(* Logix 5000 project; controller R400_500_XLS vendor 1 type 14 code 216 rev 31.11; software revision 31.01; part 24 of 32 *)
(* tags used below, declared in another part *)
   Abort1 : DINT;   // Not Used
   CycExcBuffer : UDT_CYCLE;
   Drain_RcvryTnk_with_Sump : DINT;   // 0 = Close Recovery Tank Drain Valve 1 = Open Recovery Tank Drain Valve
   DrainNo : DINT;
   DrnSmp : DINT;
   F1rinse : DINT;   // Not Used
   F2rinse : DINT;   // Not Used
   F3rinse : DINT;   // Not Used
   F4rinse : INT;   // Transition for the conductivity based evalutaion
   FINALRINSE_1 : DINT;   // Final rinse 1 id number
   FINALRINSE_9 : DINT;   // Final rinse 9 id number
   First_PwWshRnseTtr : DINT;
   Last_PwWshRnseTtr : DINT;
   M : DINT[5];   // Memory Bits
   ONS_FC13 : DINT;
   PREWASH_1 : DINT;   // Pre-wash 1 id number
   PREWASH_2 : DINT;   // Pre-wash 2 id number
   PREWASH_3 : DINT;   // Pre-wash 3 id number
   PREWASH_4 : DINT;   // Pre-wash 4 id number
   Rcvry_Tnk_Tmp : REAL;   // Water Temperature of the Heat Recovery Tank
   RINSE_1 : DINT;   // Rinse 1 id number
   RINSE_2 : DINT;   // Rinse 2 id number
   RINSE_3 : DINT;   // Rinse 3 id number
   RINSE_4 : DINT;   // Rinse 4 id number
   RLO : BOOL;   // Logic result
   Run : DINT;
   Shutdown : SINT;   // Shutdown sequence steps
   SumpWaterVolume : DINT;   // Sump Water Volume 0 =Low 1= High
   Tmr : TIMER[107];
   Trt_Drying : SINT;
   Trt_PrWsh : DINT;
   Trt_Rinse : DINT;   // Rinse steps
   Trt_Wsh : DINT;
   WASH_1 : DINT;   // Wash 1 id number
   WASH_2 : DINT;   // Wash 2 id number
   WASH_3 : DINT;   // Wash 3 id number
   WASH_4 : DINT;   // Wash 4 id number
   WASH_5 : DINT;   // Wash 5 id number
   DrainExtensionTime : DINT;
   SumpTemp : REAL;   // Sump temperature in °C
   SumpTempToCool : REAL;   // Sump temperature in °C
   TreatmentPtr : DINT;
   Unit : Hrdwre;   // Unit Configuration
(* MainProgram, continued *)

ROUTINE WSH_22_DRN_SMP_RCVR_TNK   (* ladder *)
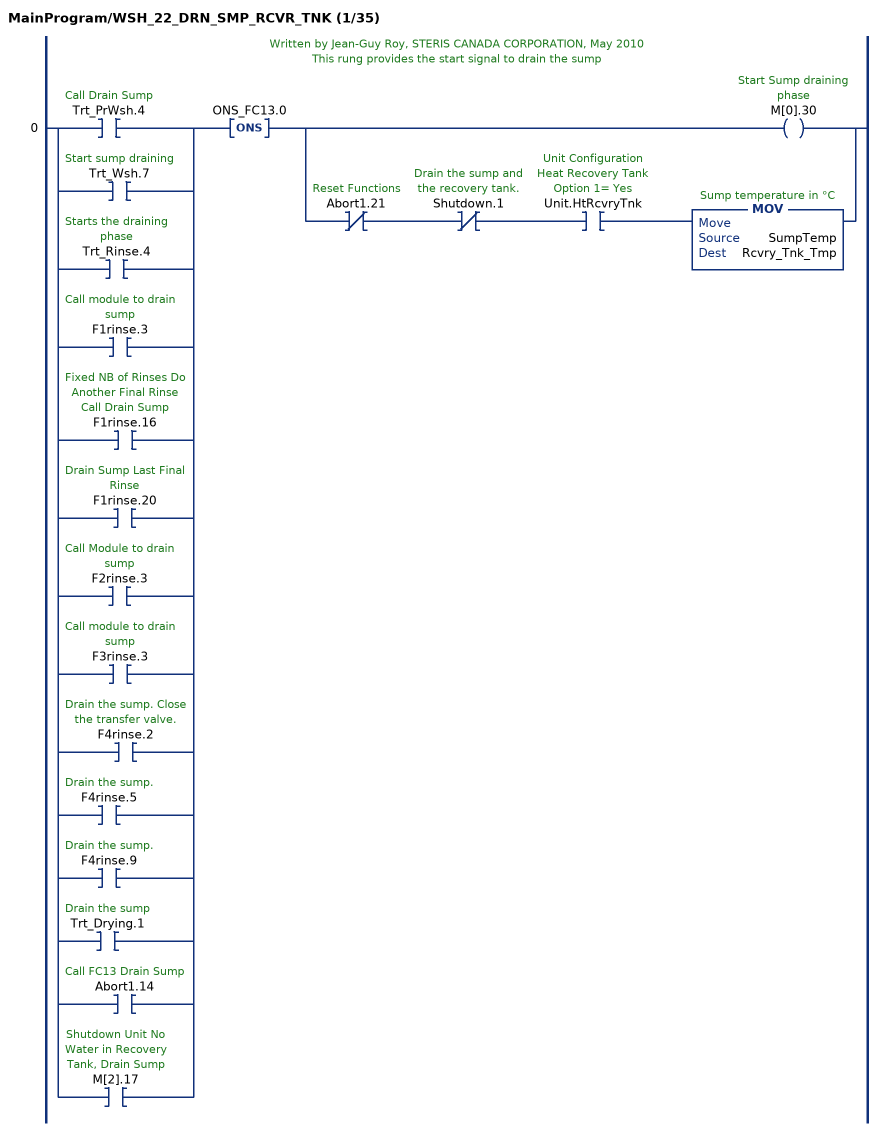
   // Written by Jean-Guy Roy, STERIS CANADA CORPORATION, May 2010
   // This rung provides the start signal to drain the sump
   0: [XIC(Trt_PrWsh.4) ,XIC(Trt_Wsh.7) ,XIC(Trt_Rinse.4) ,XIC(F1rinse.3) ,XIC(F1rinse.16) ,XIC(F1rinse.20) ,XIC(F2rinse.3) ,XIC(F3rinse.3) ,XIC(F4rinse.2) ,XIC(F4rinse.5) ,XIC(F4rinse.9) ,XIC(Trt_Drying.1) ,XIC(Abort1.14) ,XIC(M[2].17) ]ONS(ONS_FC13.0)[OTE(M[0].30) ,XIO(Abort1.21) XIO(Shutdown.1) XIC(Unit.HtRcvryTnk) MOV(SumpTemp,Rcvry_Tnk_Tmp) ];
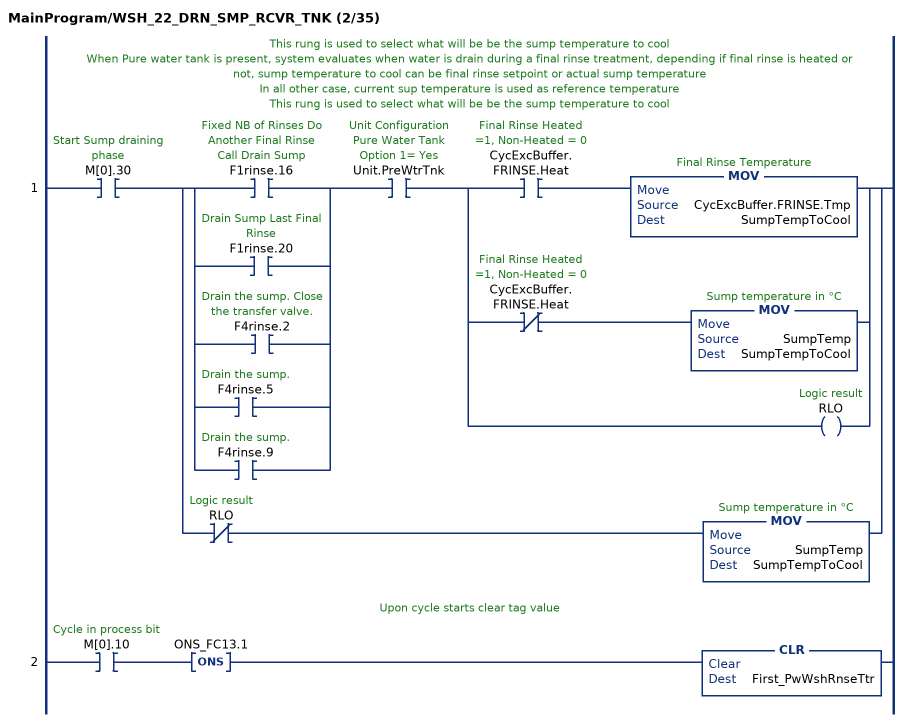
   // This rung is used to select what will be be the sump temperature to cool
   // When Pure water tank is present, system evaluates when water is drain during a final rinse treatment, depending if final rinse is heated or not, sump temperature to cool can be final rinse setpoint or actual sump temperature
   // In all other case, current sup temperature is used as reference temperature
   // This rung is used to select what will be be the sump temperature to cool
   1: XIC(M[0].30)[[XIC(F1rinse.16) ,XIC(F1rinse.20) ,XIC(F4rinse.2) ,XIC(F4rinse.5) ,XIC(F4rinse.9) ] XIC(Unit.PreWtrTnk) [XIC(CycExcBuffer.FRINSE.Heat) MOV(CycExcBuffer.FRINSE.Tmp,SumpTempToCool) ,XIO(CycExcBuffer.FRINSE.Heat) MOV(SumpTemp,SumpTempToCool) ,OTE(RLO) ] ,XIO(RLO) MOV(SumpTemp,SumpTempToCool) ];
   // Upon cycle starts clear tag value
   2: XIC(M[0].10)ONS(ONS_FC13.1)CLR(First_PwWshRnseTtr);
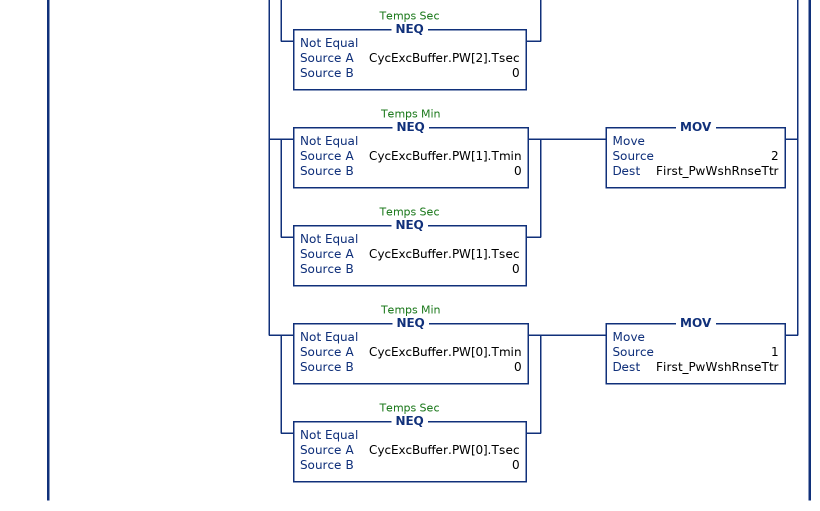
   // This rung checks which Pre-wash, Wash or Rinse treatment is the first treatment of the cycle
   // XLSV10  DGB  2018-09-17 : Added To support New Treatment
   3: XIC(M[0].10)ONS(ONS_FC13.2)[[NEQ(CycExcBuffer.RINSE[3].Tmin,0) ,NEQ(CycExcBuffer.RINSE[3].Tsec,0) ] MOV(13,First_PwWshRnseTtr) ,[NEQ(CycExcBuffer.RINSE[2].Tmin,0) ,NEQ(CycExcBuffer.RINSE[2].Tsec,0) ] MOV(12,First_PwWshRnseTtr) ,[NEQ(CycExcBuffer.RINSE[1].Tmin,0) ,NEQ(CycExcBuffer.RINSE[1].Tsec,0) ] MOV(11,First_PwWshRnseTtr) ,[NEQ(CycExcBuffer.RINSE[0].Tmin,0) ,NEQ(CycExcBuffer.RINSE[0].Tsec,0) ] MOV(10,First_PwWshRnseTtr) ,[NEQ(CycExcBuffer.WSH[4].Tmin,0) ,NEQ(CycExcBuffer.WSH[4].Tsec,0) ] MOV(9,First_PwWshRnseTtr) ,[NEQ(CycExcBuffer.WSH[3].Tmin,0) ,NEQ(CycExcBuffer.WSH[3].Tsec,0) ] MOV(8,First_PwWshRnseTtr) ,[NEQ(CycExcBuffer.WSH[2].Tmin,0) ,NEQ(CycExcBuffer.WSH[2].Tsec,0) ] MOV(7,First_PwWshRnseTtr) ,[NEQ(CycExcBuffer.WSH[1].Tmin,0) ,NEQ(CycExcBuffer.WSH[1].Tsec,0) ] MOV(6,First_PwWshRnseTtr) ,[NEQ(CycExcBuffer.WSH[0].Tmin,0) ,NEQ(CycExcBuffer.WSH[0].Tsec,0) ] MOV(5,First_PwWshRnseTtr) ,[NEQ(CycExcBuffer.PW[3].Tmin,0) ,NEQ(CycExcBuffer.PW[3].Tsec,0) ] MOV(4,First_PwWshRnseTtr) ,[NEQ(CycExcBuffer.PW[2].Tmin,0) ,NEQ(CycExcBuffer.PW[2].Tsec,0) ] MOV(3,First_PwWshRnseTtr) ,[NEQ(CycExcBuffer.PW[1].Tmin,0) ,NEQ(CycExcBuffer.PW[1].Tsec,0) ] MOV(2,First_PwWshRnseTtr) ,[NEQ(CycExcBuffer.PW[0].Tmin,0) ,NEQ(CycExcBuffer.PW[0].Tsec,0) ] MOV(1,First_PwWshRnseTtr) ];
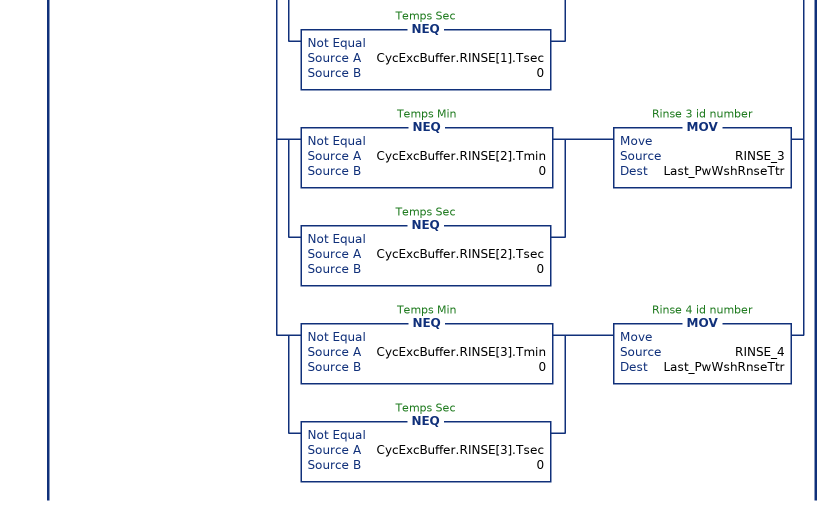
   // This rung detect which recirculated treatment is the last treatment of the cycle
   // XLSV10  DGB  2018-09-07 : Modified to support Added Treatments
   4: XIC(M[0].10)ONS(ONS_FC13.10)[[NEQ(CycExcBuffer.PW[0].Tmin,0) ,NEQ(CycExcBuffer.PW[0].Tsec,0) ] MOV(PREWASH_1,Last_PwWshRnseTtr) ,[NEQ(CycExcBuffer.PW[1].Tmin,0) ,NEQ(CycExcBuffer.PW[1].Tsec,0) ] MOV(PREWASH_2,Last_PwWshRnseTtr) ,[NEQ(CycExcBuffer.PW[2].Tmin,0) ,NEQ(CycExcBuffer.PW[2].Tsec,0) ] MOV(PREWASH_3,Last_PwWshRnseTtr) ,[NEQ(CycExcBuffer.PW[3].Tmin,0) ,NEQ(CycExcBuffer.PW[3].Tsec,0) ] MOV(PREWASH_4,Last_PwWshRnseTtr) ,[NEQ(CycExcBuffer.WSH[0].Tmin,0) ,NEQ(CycExcBuffer.WSH[0].Tsec,0) ] MOV(WASH_1,Last_PwWshRnseTtr) ,[NEQ(CycExcBuffer.WSH[1].Tmin,0) ,NEQ(CycExcBuffer.WSH[1].Tsec,0) ] MOV(WASH_2,Last_PwWshRnseTtr) ,[NEQ(CycExcBuffer.WSH[2].Tmin,0) ,NEQ(CycExcBuffer.WSH[2].Tsec,0) ] MOV(WASH_3,Last_PwWshRnseTtr) ,[NEQ(CycExcBuffer.WSH[3].Tmin,0) ,NEQ(CycExcBuffer.WSH[3].Tsec,0) ] MOV(WASH_4,Last_PwWshRnseTtr) ,[NEQ(CycExcBuffer.WSH[4].Tmin,0) ,NEQ(CycExcBuffer.WSH[4].Tsec,0) ] MOV(WASH_5,Last_PwWshRnseTtr) ,[NEQ(CycExcBuffer.RINSE[0].Tmin,0) ,NEQ(CycExcBuffer.RINSE[0].Tsec,0) ] MOV(RINSE_1,Last_PwWshRnseTtr) ,[NEQ(CycExcBuffer.RINSE[1].Tmin,0) ,NEQ(CycExcBuffer.RINSE[1].Tsec,0) ] MOV(RINSE_2,Last_PwWshRnseTtr) ,[NEQ(CycExcBuffer.RINSE[2].Tmin,0) ,NEQ(CycExcBuffer.RINSE[2].Tsec,0) ] MOV(RINSE_3,Last_PwWshRnseTtr) ,[NEQ(CycExcBuffer.RINSE[3].Tmin,0) ,NEQ(CycExcBuffer.RINSE[3].Tsec,0) ] MOV(RINSE_4,Last_PwWshRnseTtr) ];
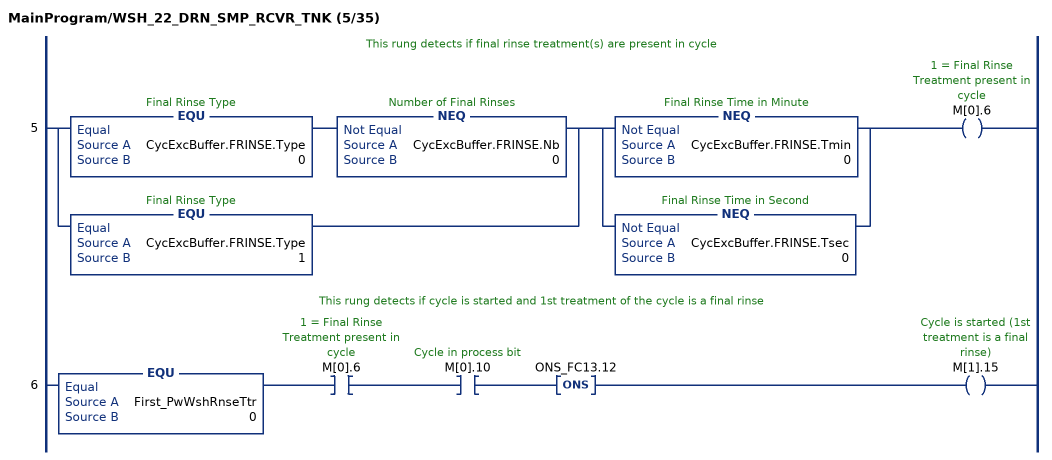
   // This rung detects if final rinse treatment(s) are present in cycle
   5: [EQU(CycExcBuffer.FRINSE.Type,0) NEQ(CycExcBuffer.FRINSE.Nb,0) ,EQU(CycExcBuffer.FRINSE.Type,1) ][NEQ(CycExcBuffer.FRINSE.Tmin,0) ,NEQ(CycExcBuffer.FRINSE.Tsec,0) ]OTE(M[0].6);
   // This rung detects if cycle is started and 1st treatment of the cycle is a final rinse
   6: EQU(First_PwWshRnseTtr,0)XIC(M[0].6)XIC(M[0].10)ONS(ONS_FC13.12)OTE(M[1].15);
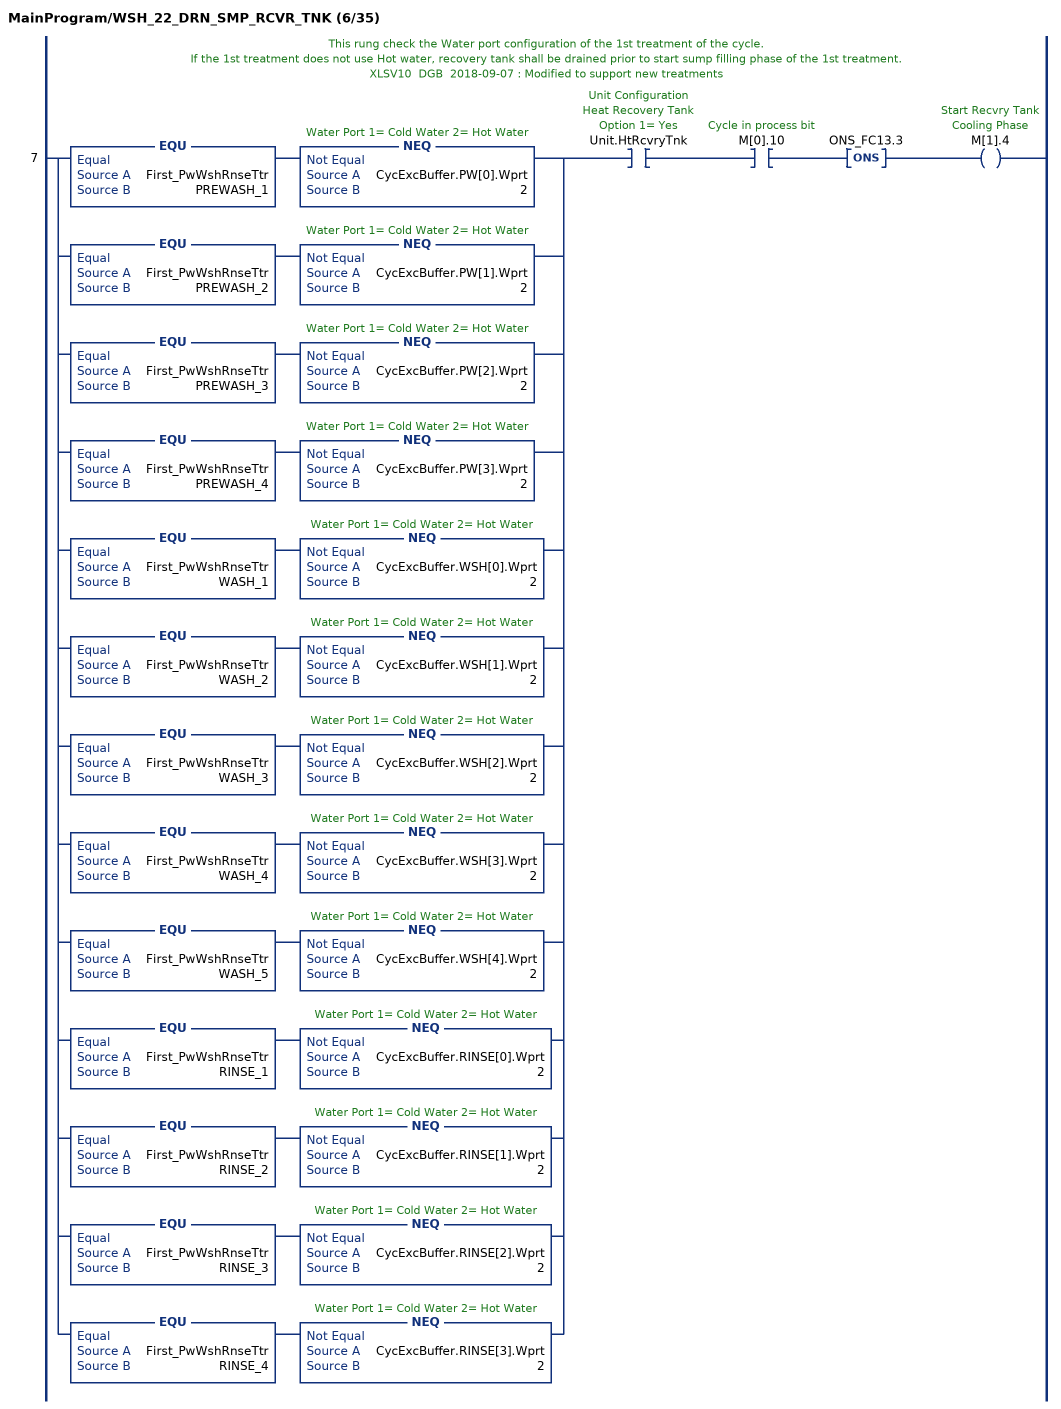
   // This rung check the Water port configuration of the 1st treatment of the cycle.
   // If the 1st treatment does not use Hot water, recovery tank shall be drained prior to start sump filling phase of the 1st treatment.
   // XLSV10  DGB  2018-09-07 : Modified to support new treatments
   7: [EQU(First_PwWshRnseTtr,PREWASH_1) NEQ(CycExcBuffer.PW[0].Wprt,2) ,EQU(First_PwWshRnseTtr,PREWASH_2) NEQ(CycExcBuffer.PW[1].Wprt,2) ,EQU(First_PwWshRnseTtr,PREWASH_3) NEQ(CycExcBuffer.PW[2].Wprt,2) ,EQU(First_PwWshRnseTtr,PREWASH_4) NEQ(CycExcBuffer.PW[3].Wprt,2) ,EQU(First_PwWshRnseTtr,WASH_1) NEQ(CycExcBuffer.WSH[0].Wprt,2) ,EQU(First_PwWshRnseTtr,WASH_2) NEQ(CycExcBuffer.WSH[1].Wprt,2) ,EQU(First_PwWshRnseTtr,WASH_3) NEQ(CycExcBuffer.WSH[2].Wprt,2) ,EQU(First_PwWshRnseTtr,WASH_4) NEQ(CycExcBuffer.WSH[3].Wprt,2) ,EQU(First_PwWshRnseTtr,WASH_5) NEQ(CycExcBuffer.WSH[4].Wprt,2) ,EQU(First_PwWshRnseTtr,RINSE_1) NEQ(CycExcBuffer.RINSE[0].Wprt,2) ,EQU(First_PwWshRnseTtr,RINSE_2) NEQ(CycExcBuffer.RINSE[1].Wprt,2) ,EQU(First_PwWshRnseTtr,RINSE_3) NEQ(CycExcBuffer.RINSE[2].Wprt,2) ,EQU(First_PwWshRnseTtr,RINSE_4) NEQ(CycExcBuffer.RINSE[3].Wprt,2) ]XIC(Unit.HtRcvryTnk)XIC(M[0].10)ONS(ONS_FC13.3)OTE(M[1].4);
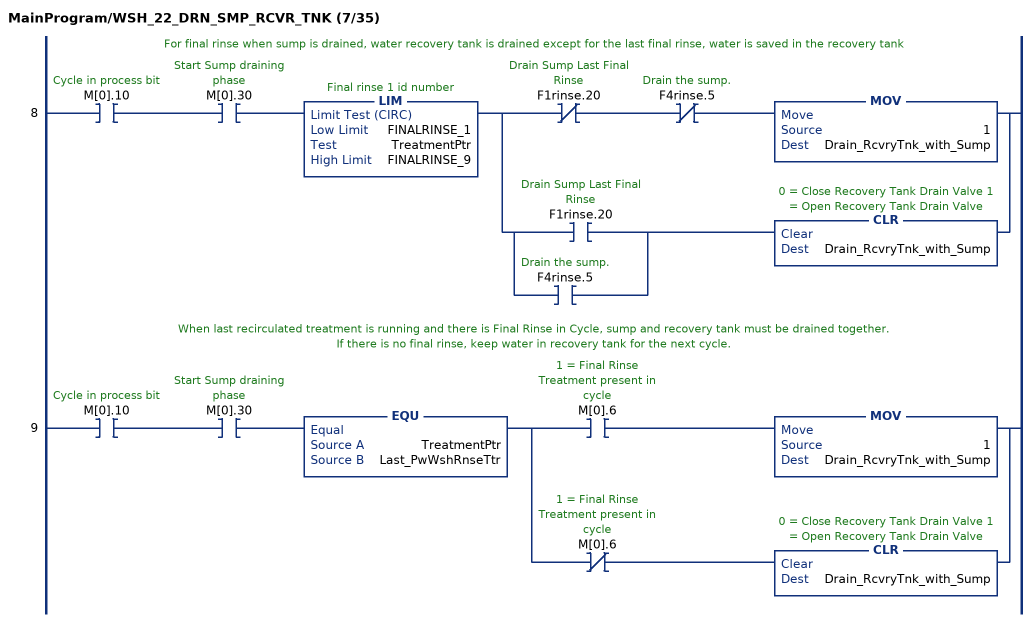
   // For final rinse when sump is drained, water recovery tank is drained except for the last final rinse, water is saved in the recovery tank
   8: XIC(M[0].10)XIC(M[0].30)LIM(FINALRINSE_1,TreatmentPtr,FINALRINSE_9)[XIO(F1rinse.20) XIO(F4rinse.5) MOV(1,Drain_RcvryTnk_with_Sump) ,[XIC(F1rinse.20) ,XIC(F4rinse.5) ] CLR(Drain_RcvryTnk_with_Sump) ];
   // When last recirculated treatment is running and there is Final Rinse in Cycle, sump and recovery tank must be drained together.
   // If there is no final rinse, keep water in recovery tank for the next cycle.
   9: XIC(M[0].10)XIC(M[0].30)EQU(TreatmentPtr,Last_PwWshRnseTtr)[XIC(M[0].6) MOV(1,Drain_RcvryTnk_with_Sump) ,XIO(M[0].6) CLR(Drain_RcvryTnk_with_Sump) ];
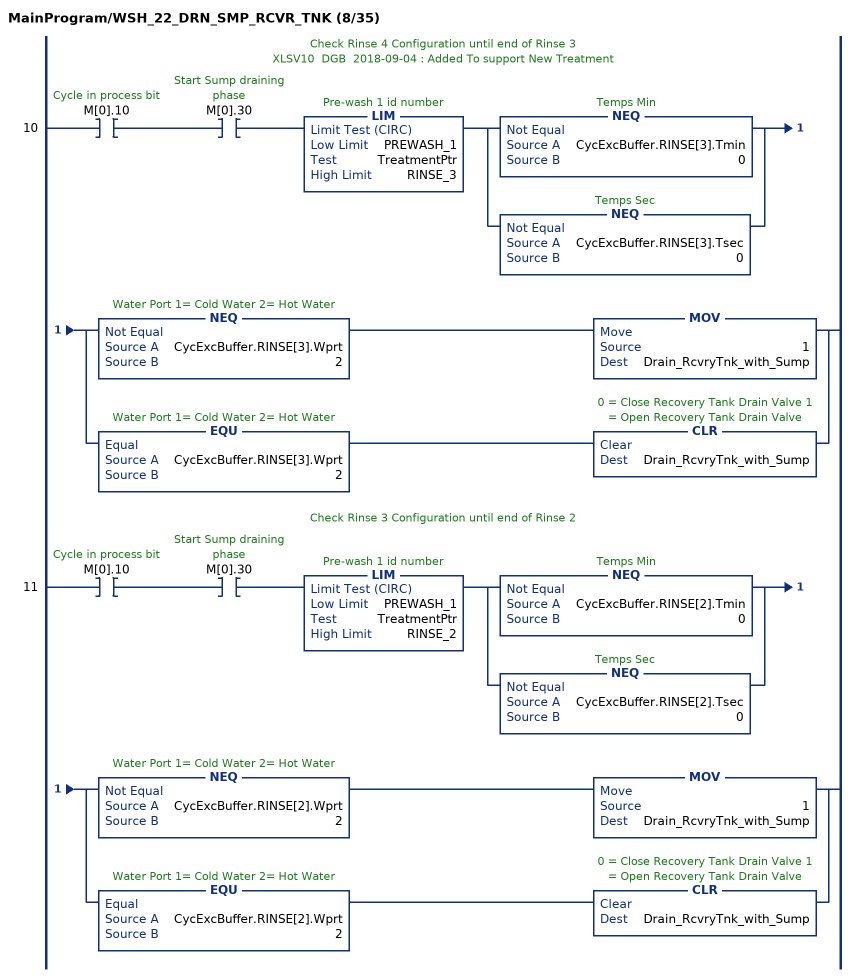
   // Check Rinse 4 Configuration until end of Rinse 3
   // XLSV10  DGB  2018-09-04 : Added To support New Treatment
   10: XIC(M[0].10)XIC(M[0].30)LIM(PREWASH_1,TreatmentPtr,RINSE_3)[NEQ(CycExcBuffer.RINSE[3].Tmin,0) ,NEQ(CycExcBuffer.RINSE[3].Tsec,0) ][NEQ(CycExcBuffer.RINSE[3].Wprt,2) MOV(1,Drain_RcvryTnk_with_Sump) ,EQU(CycExcBuffer.RINSE[3].Wprt,2) CLR(Drain_RcvryTnk_with_Sump) ];
   // Check Rinse 3 Configuration until end of Rinse 2
   11: XIC(M[0].10)XIC(M[0].30)LIM(PREWASH_1,TreatmentPtr,RINSE_2)[NEQ(CycExcBuffer.RINSE[2].Tmin,0) ,NEQ(CycExcBuffer.RINSE[2].Tsec,0) ][NEQ(CycExcBuffer.RINSE[2].Wprt,2) MOV(1,Drain_RcvryTnk_with_Sump) ,EQU(CycExcBuffer.RINSE[2].Wprt,2) CLR(Drain_RcvryTnk_with_Sump) ];
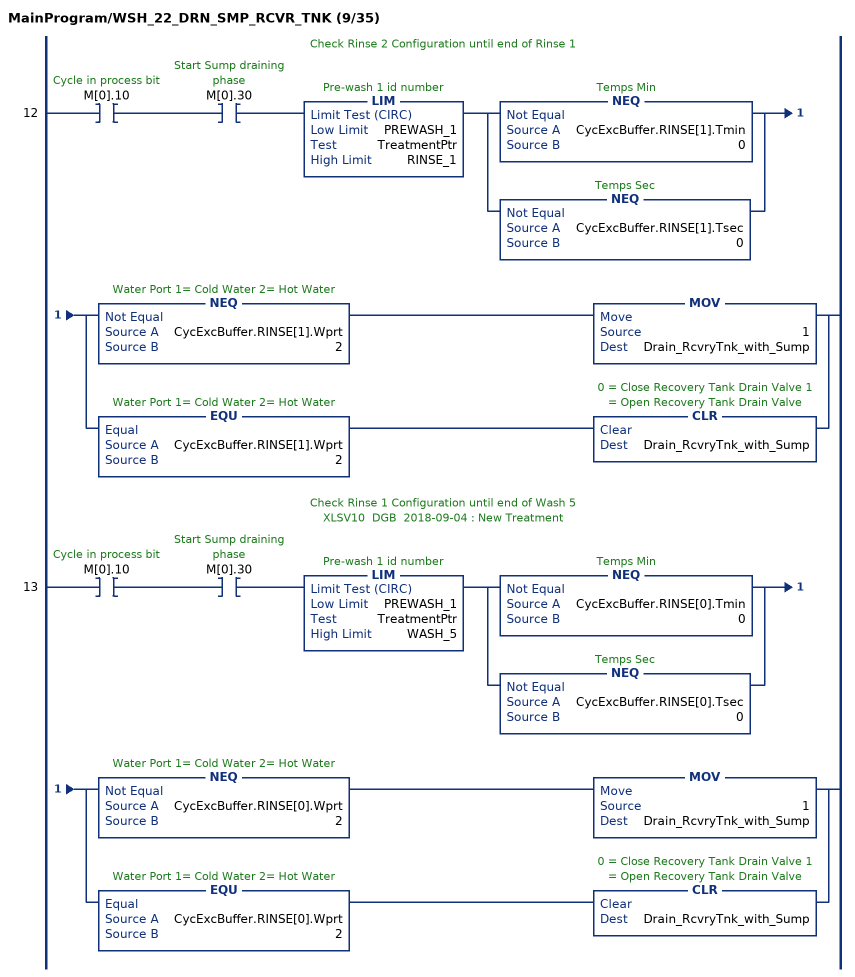
   // Check Rinse 2 Configuration until end of Rinse 1
   12: XIC(M[0].10)XIC(M[0].30)LIM(PREWASH_1,TreatmentPtr,RINSE_1)[NEQ(CycExcBuffer.RINSE[1].Tmin,0) ,NEQ(CycExcBuffer.RINSE[1].Tsec,0) ][NEQ(CycExcBuffer.RINSE[1].Wprt,2) MOV(1,Drain_RcvryTnk_with_Sump) ,EQU(CycExcBuffer.RINSE[1].Wprt,2) CLR(Drain_RcvryTnk_with_Sump) ];
   // Check Rinse 1 Configuration until end of Wash 5
   // XLSV10  DGB  2018-09-04 : New Treatment
   13: XIC(M[0].10)XIC(M[0].30)LIM(PREWASH_1,TreatmentPtr,WASH_5)[NEQ(CycExcBuffer.RINSE[0].Tmin,0) ,NEQ(CycExcBuffer.RINSE[0].Tsec,0) ][NEQ(CycExcBuffer.RINSE[0].Wprt,2) MOV(1,Drain_RcvryTnk_with_Sump) ,EQU(CycExcBuffer.RINSE[0].Wprt,2) CLR(Drain_RcvryTnk_with_Sump) ];
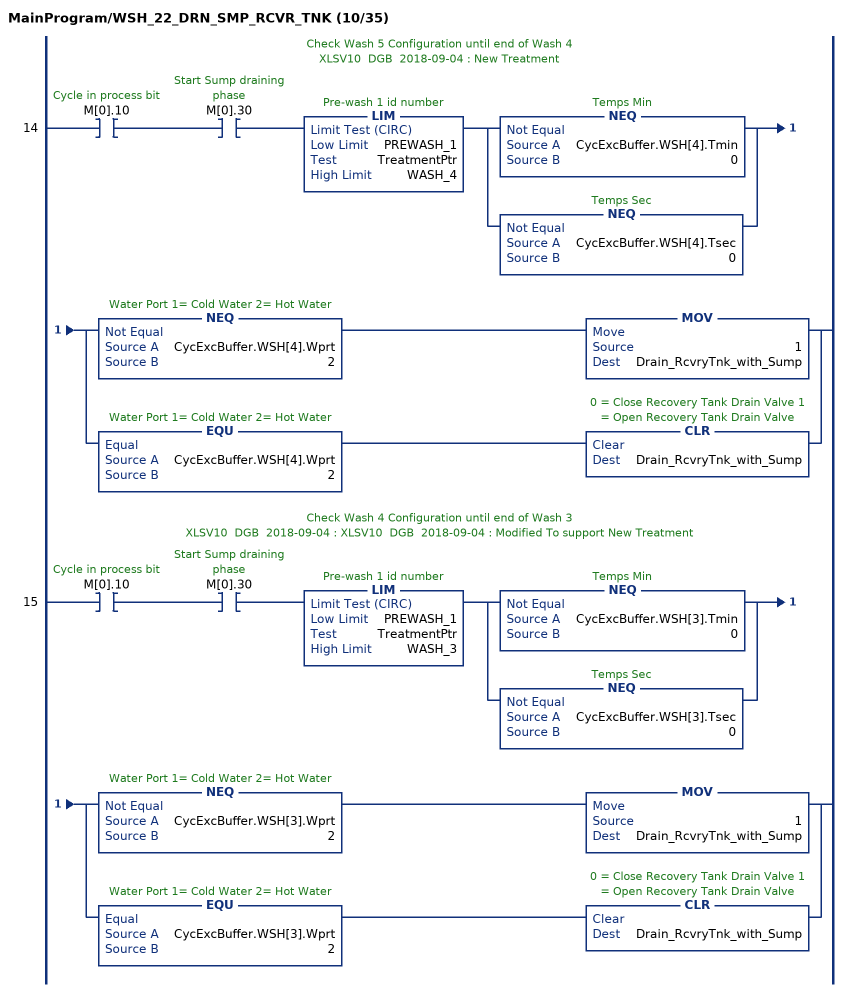
   // Check Wash 5 Configuration until end of Wash 4
   // XLSV10  DGB  2018-09-04 : New Treatment
   14: XIC(M[0].10)XIC(M[0].30)LIM(PREWASH_1,TreatmentPtr,WASH_4)[NEQ(CycExcBuffer.WSH[4].Tmin,0) ,NEQ(CycExcBuffer.WSH[4].Tsec,0) ][NEQ(CycExcBuffer.WSH[4].Wprt,2) MOV(1,Drain_RcvryTnk_with_Sump) ,EQU(CycExcBuffer.WSH[4].Wprt,2) CLR(Drain_RcvryTnk_with_Sump) ];
   // Check Wash 4 Configuration until end of Wash 3
   // XLSV10  DGB  2018-09-04 : XLSV10  DGB  2018-09-04 : Modified To support New Treatment
   15: XIC(M[0].10)XIC(M[0].30)LIM(PREWASH_1,TreatmentPtr,WASH_3)[NEQ(CycExcBuffer.WSH[3].Tmin,0) ,NEQ(CycExcBuffer.WSH[3].Tsec,0) ][NEQ(CycExcBuffer.WSH[3].Wprt,2) MOV(1,Drain_RcvryTnk_with_Sump) ,EQU(CycExcBuffer.WSH[3].Wprt,2) CLR(Drain_RcvryTnk_with_Sump) ];
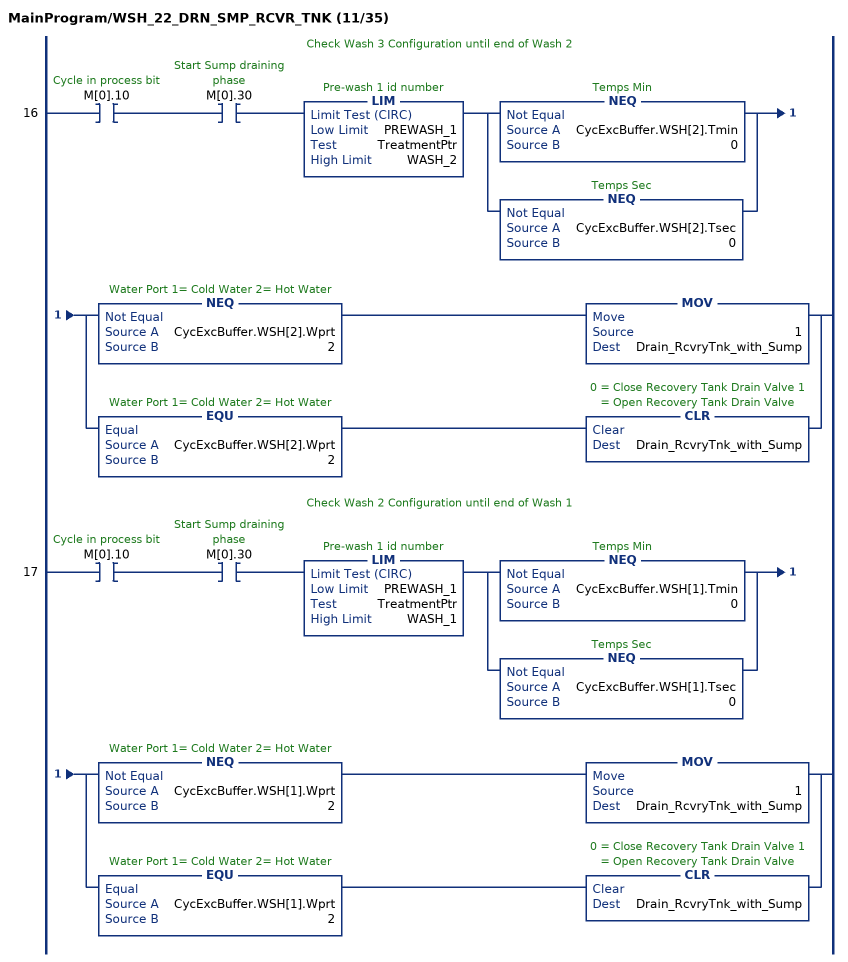
   // Check Wash 3 Configuration until end of Wash 2
   16: XIC(M[0].10)XIC(M[0].30)LIM(PREWASH_1,TreatmentPtr,WASH_2)[NEQ(CycExcBuffer.WSH[2].Tmin,0) ,NEQ(CycExcBuffer.WSH[2].Tsec,0) ][NEQ(CycExcBuffer.WSH[2].Wprt,2) MOV(1,Drain_RcvryTnk_with_Sump) ,EQU(CycExcBuffer.WSH[2].Wprt,2) CLR(Drain_RcvryTnk_with_Sump) ];
   // Check Wash 2 Configuration until end of Wash 1
   17: XIC(M[0].10)XIC(M[0].30)LIM(PREWASH_1,TreatmentPtr,WASH_1)[NEQ(CycExcBuffer.WSH[1].Tmin,0) ,NEQ(CycExcBuffer.WSH[1].Tsec,0) ][NEQ(CycExcBuffer.WSH[1].Wprt,2) MOV(1,Drain_RcvryTnk_with_Sump) ,EQU(CycExcBuffer.WSH[1].Wprt,2) CLR(Drain_RcvryTnk_with_Sump) ];
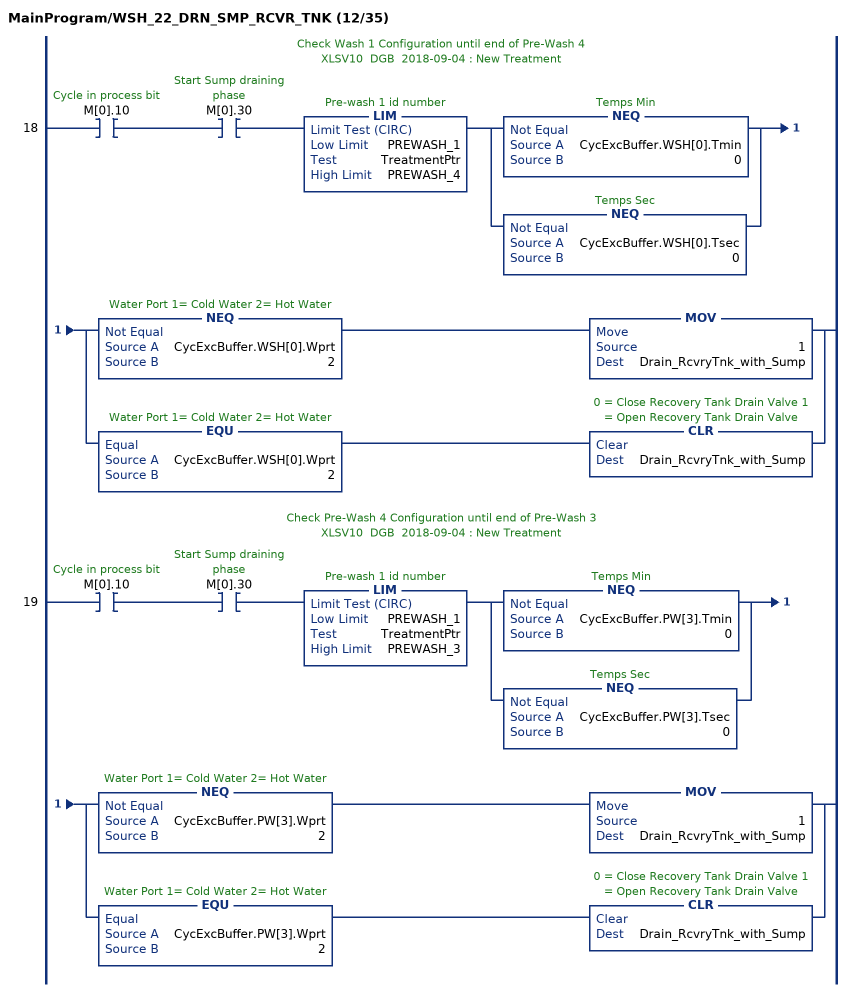
   // Check Wash 1 Configuration until end of Pre-Wash 4
   // XLSV10  DGB  2018-09-04 : New Treatment
   18: XIC(M[0].10)XIC(M[0].30)LIM(PREWASH_1,TreatmentPtr,PREWASH_4)[NEQ(CycExcBuffer.WSH[0].Tmin,0) ,NEQ(CycExcBuffer.WSH[0].Tsec,0) ][NEQ(CycExcBuffer.WSH[0].Wprt,2) MOV(1,Drain_RcvryTnk_with_Sump) ,EQU(CycExcBuffer.WSH[0].Wprt,2) CLR(Drain_RcvryTnk_with_Sump) ];
   // Check Pre-Wash 4 Configuration until end of Pre-Wash 3
   // XLSV10  DGB  2018-09-04 : New Treatment
   19: XIC(M[0].10)XIC(M[0].30)LIM(PREWASH_1,TreatmentPtr,PREWASH_3)[NEQ(CycExcBuffer.PW[3].Tmin,0) ,NEQ(CycExcBuffer.PW[3].Tsec,0) ][NEQ(CycExcBuffer.PW[3].Wprt,2) MOV(1,Drain_RcvryTnk_with_Sump) ,EQU(CycExcBuffer.PW[3].Wprt,2) CLR(Drain_RcvryTnk_with_Sump) ];
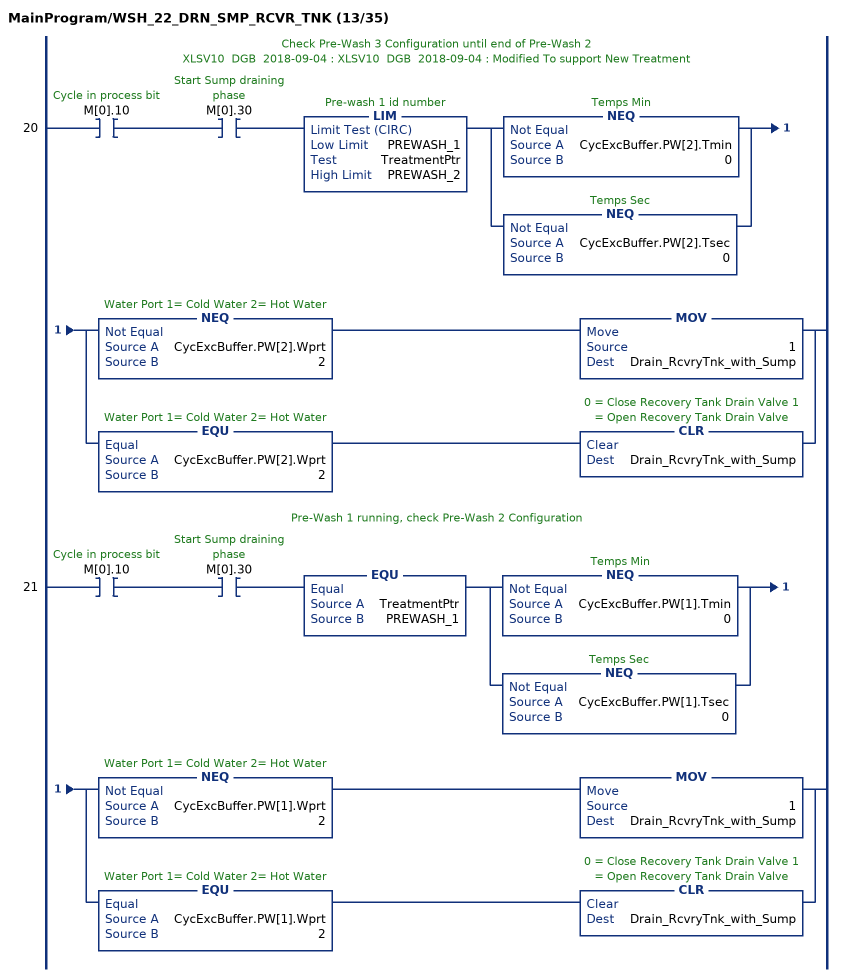
   // Check Pre-Wash 3 Configuration until end of Pre-Wash 2
   // XLSV10  DGB  2018-09-04 : XLSV10  DGB  2018-09-04 : Modified To support New Treatment
   20: XIC(M[0].10)XIC(M[0].30)LIM(PREWASH_1,TreatmentPtr,PREWASH_2)[NEQ(CycExcBuffer.PW[2].Tmin,0) ,NEQ(CycExcBuffer.PW[2].Tsec,0) ][NEQ(CycExcBuffer.PW[2].Wprt,2) MOV(1,Drain_RcvryTnk_with_Sump) ,EQU(CycExcBuffer.PW[2].Wprt,2) CLR(Drain_RcvryTnk_with_Sump) ];
   // Pre-Wash 1 running, check Pre-Wash 2 Configuration
   21: XIC(M[0].10)XIC(M[0].30)EQU(TreatmentPtr,PREWASH_1)[NEQ(CycExcBuffer.PW[1].Tmin,0) ,NEQ(CycExcBuffer.PW[1].Tsec,0) ][NEQ(CycExcBuffer.PW[1].Wprt,2) MOV(1,Drain_RcvryTnk_with_Sump) ,EQU(CycExcBuffer.PW[1].Wprt,2) CLR(Drain_RcvryTnk_with_Sump) ];
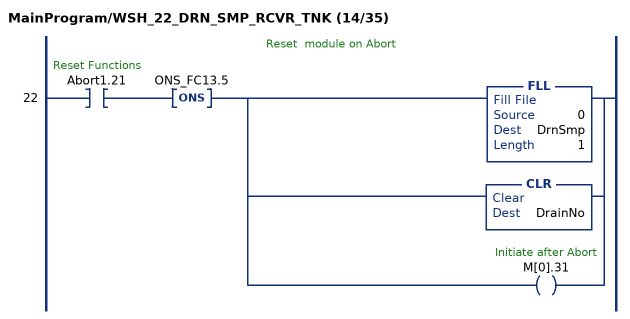
   // Reset  module on Abort
   22: XIC(Abort1.21)ONS(ONS_FC13.5)[FLL(0,DrnSmp,1) ,CLR(DrainNo) ,OTE(M[0].31) ];
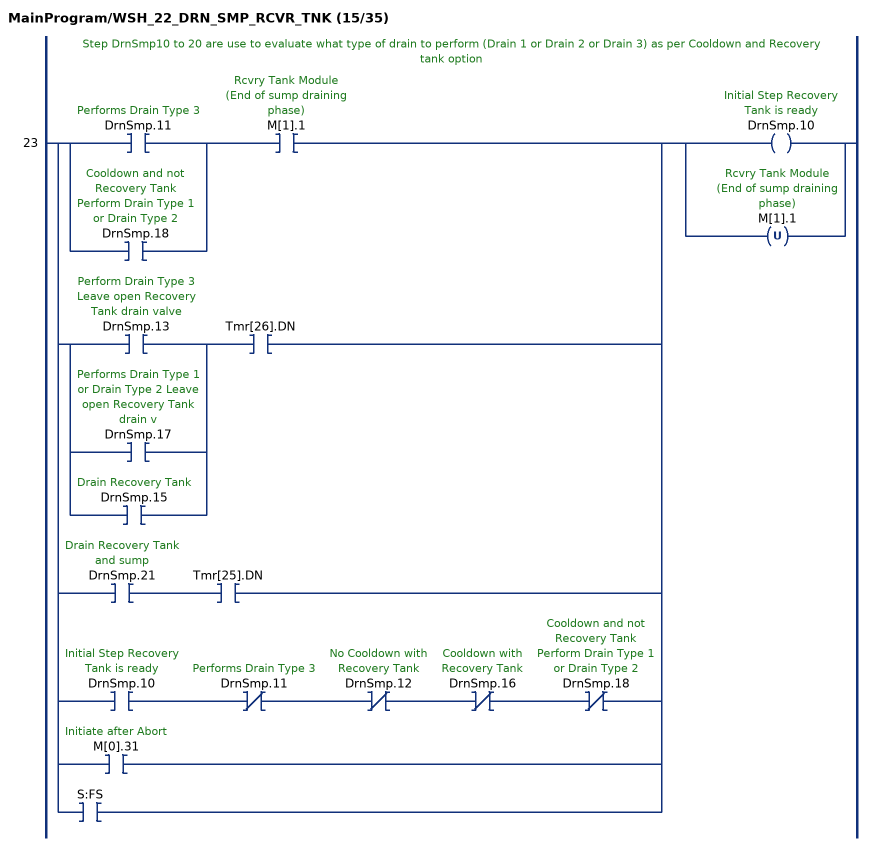
   // Step DrnSmp10 to 20 are use to evaluate what type of drain to perform (Drain 1 or Drain 2 or Drain 3) as per Cooldown and Recovery tank option
   23: [[[XIC(DrnSmp.11) ,XIC(DrnSmp.18) ] XIC(M[1].1) ,[XIC(DrnSmp.13) ,XIC(DrnSmp.17) ,XIC(DrnSmp.15) ] XIC(Tmr[26].DN) ,XIC(DrnSmp.21) XIC(Tmr[25].DN) ] ,XIC(DrnSmp.10) XIO(DrnSmp.11) XIO(DrnSmp.12) XIO(DrnSmp.16) XIO(DrnSmp.18) ,XIC(M[0].31) ,XIC(S:FS) ][OTE(DrnSmp.10) ,OTU(M[1].1) ];
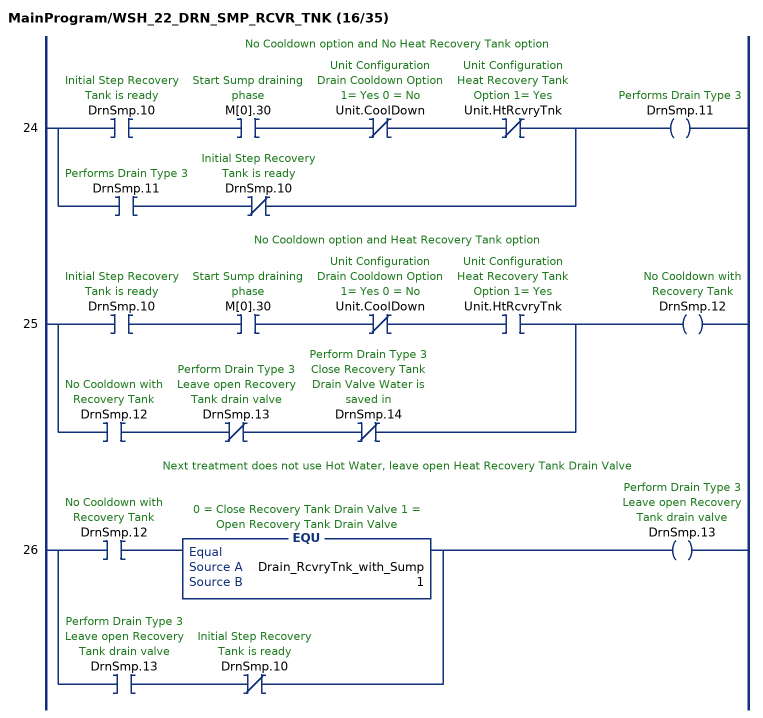
   // No Cooldown option and No Heat Recovery Tank option
   24: [XIC(DrnSmp.10) XIC(M[0].30) XIO(Unit.CoolDown) XIO(Unit.HtRcvryTnk) ,XIC(DrnSmp.11) XIO(DrnSmp.10) ]OTE(DrnSmp.11);
   // No Cooldown option and Heat Recovery Tank option
   25: [XIC(DrnSmp.10) XIC(M[0].30) XIO(Unit.CoolDown) XIC(Unit.HtRcvryTnk) ,XIC(DrnSmp.12) XIO(DrnSmp.13) XIO(DrnSmp.14) ]OTE(DrnSmp.12);
   // Next treatment does not use Hot Water, leave open Heat Recovery Tank Drain Valve
   26: [XIC(DrnSmp.12) EQU(Drain_RcvryTnk_with_Sump,1) ,XIC(DrnSmp.13) XIO(DrnSmp.10) ]OTE(DrnSmp.13);
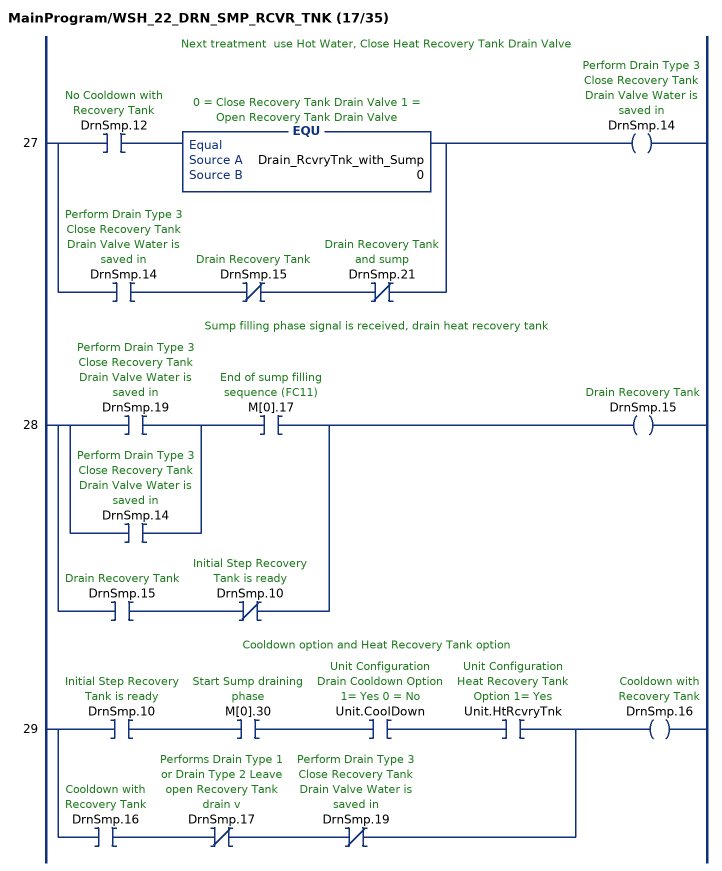
   // Next treatment  use Hot Water, Close Heat Recovery Tank Drain Valve
   27: [XIC(DrnSmp.12) EQU(Drain_RcvryTnk_with_Sump,0) ,XIC(DrnSmp.14) XIO(DrnSmp.15) XIO(DrnSmp.21) ]OTE(DrnSmp.14);
   // Sump filling phase signal is received, drain heat recovery tank
   28: [[XIC(DrnSmp.19) ,XIC(DrnSmp.14) ] XIC(M[0].17) ,XIC(DrnSmp.15) XIO(DrnSmp.10) ]OTE(DrnSmp.15);
   // Cooldown option and Heat Recovery Tank option
   29: [XIC(DrnSmp.10) XIC(M[0].30) XIC(Unit.CoolDown) XIC(Unit.HtRcvryTnk) ,XIC(DrnSmp.16) XIO(DrnSmp.17) XIO(DrnSmp.19) ]OTE(DrnSmp.16);
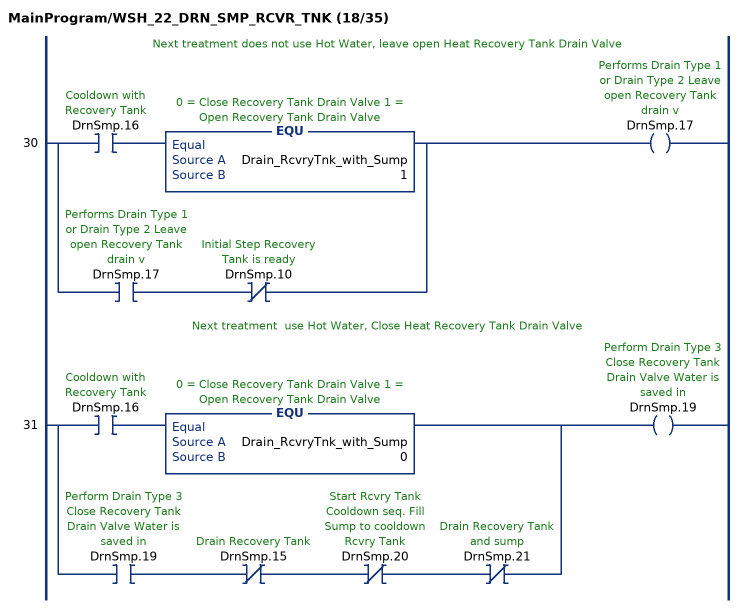
   // Next treatment does not use Hot Water, leave open Heat Recovery Tank Drain Valve
   30: [XIC(DrnSmp.16) EQU(Drain_RcvryTnk_with_Sump,1) ,XIC(DrnSmp.17) XIO(DrnSmp.10) ]OTE(DrnSmp.17);
   // Next treatment  use Hot Water, Close Heat Recovery Tank Drain Valve
   31: [XIC(DrnSmp.16) EQU(Drain_RcvryTnk_with_Sump,0) ,XIC(DrnSmp.19) XIO(DrnSmp.15) XIO(DrnSmp.20) XIO(DrnSmp.21) ]OTE(DrnSmp.19);
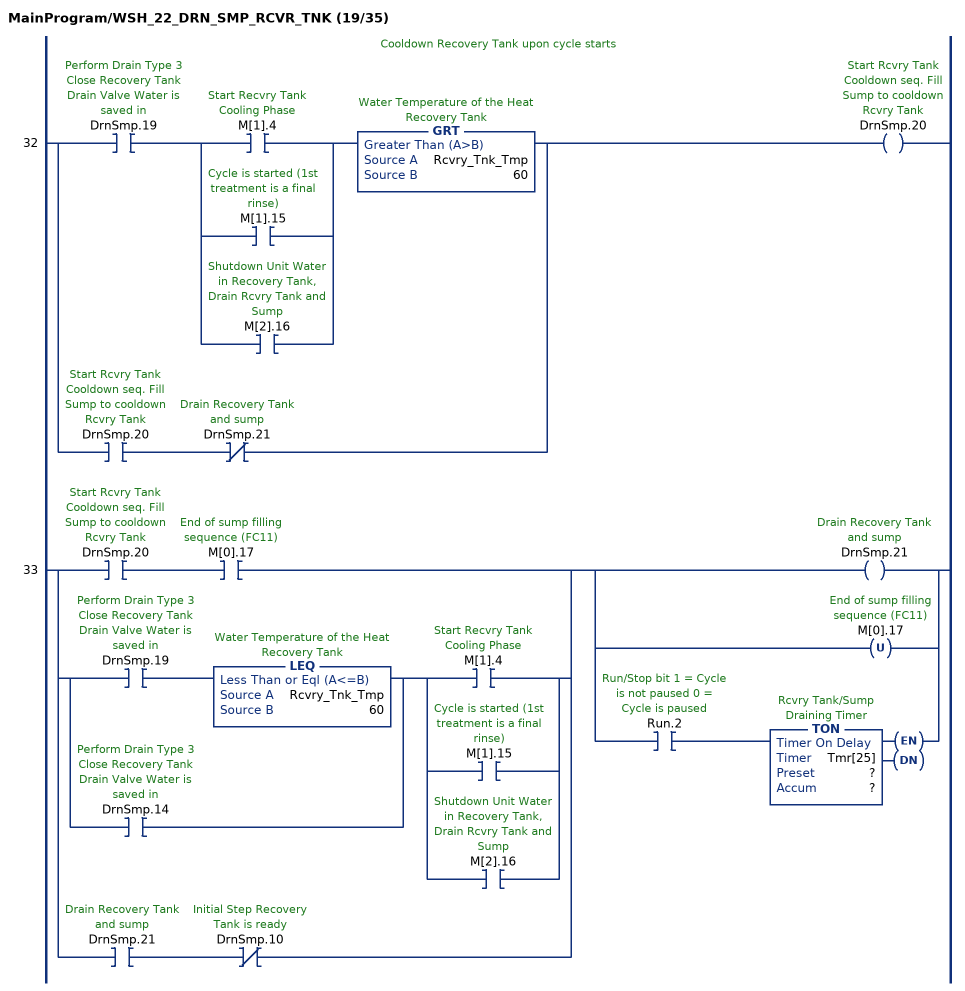
   // Cooldown Recovery Tank upon cycle starts
   32: [XIC(DrnSmp.19) [XIC(M[1].4) ,XIC(M[1].15) ,XIC(M[2].16) ] GRT(Rcvry_Tnk_Tmp,60) ,XIC(DrnSmp.20) XIO(DrnSmp.21) ]OTE(DrnSmp.20);
   33: [XIC(DrnSmp.20) XIC(M[0].17) ,[XIC(DrnSmp.19) LEQ(Rcvry_Tnk_Tmp,60) ,XIC(DrnSmp.14) ] [XIC(M[1].4) ,XIC(M[1].15) ,XIC(M[2].16) ] ,XIC(DrnSmp.21) XIO(DrnSmp.10) ][OTE(DrnSmp.21) ,OTU(M[0].17) ,XIC(Run.2) TON(Tmr[25],?,?) ];
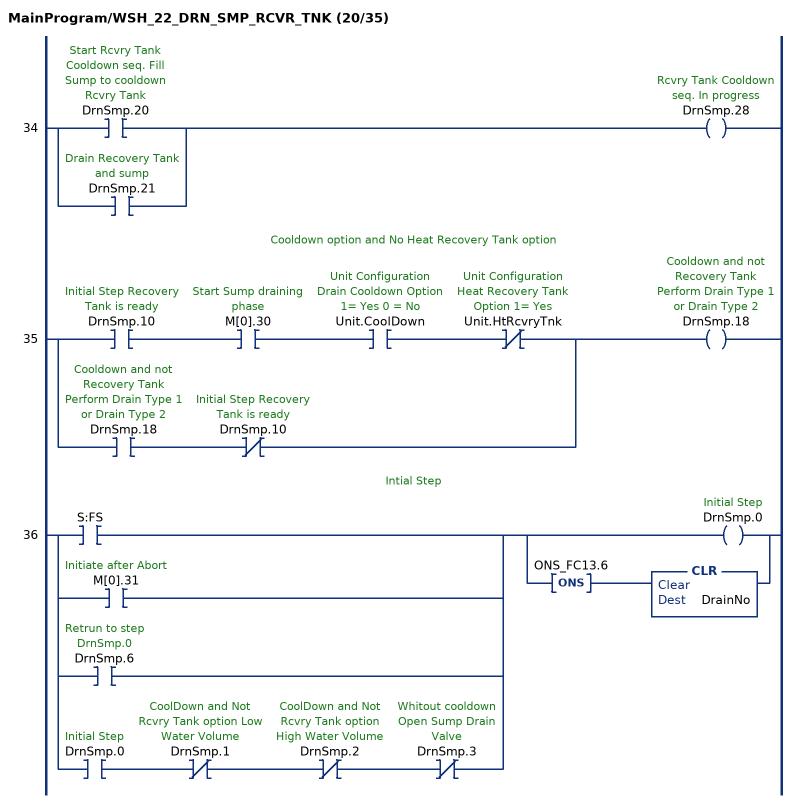
   34: [XIC(DrnSmp.20) ,XIC(DrnSmp.21) ]OTE(DrnSmp.28);
   // Cooldown option and No Heat Recovery Tank option
   35: [XIC(DrnSmp.10) XIC(M[0].30) XIC(Unit.CoolDown) XIO(Unit.HtRcvryTnk) ,XIC(DrnSmp.18) XIO(DrnSmp.10) ]OTE(DrnSmp.18);
   // Intial Step
   36: [XIC(S:FS) ,XIC(M[0].31) ,XIC(DrnSmp.6) ,XIC(DrnSmp.0) XIO(DrnSmp.1) XIO(DrnSmp.2) XIO(DrnSmp.3) ][OTE(DrnSmp.0) ,ONS(ONS_FC13.6) CLR(DrainNo) ];
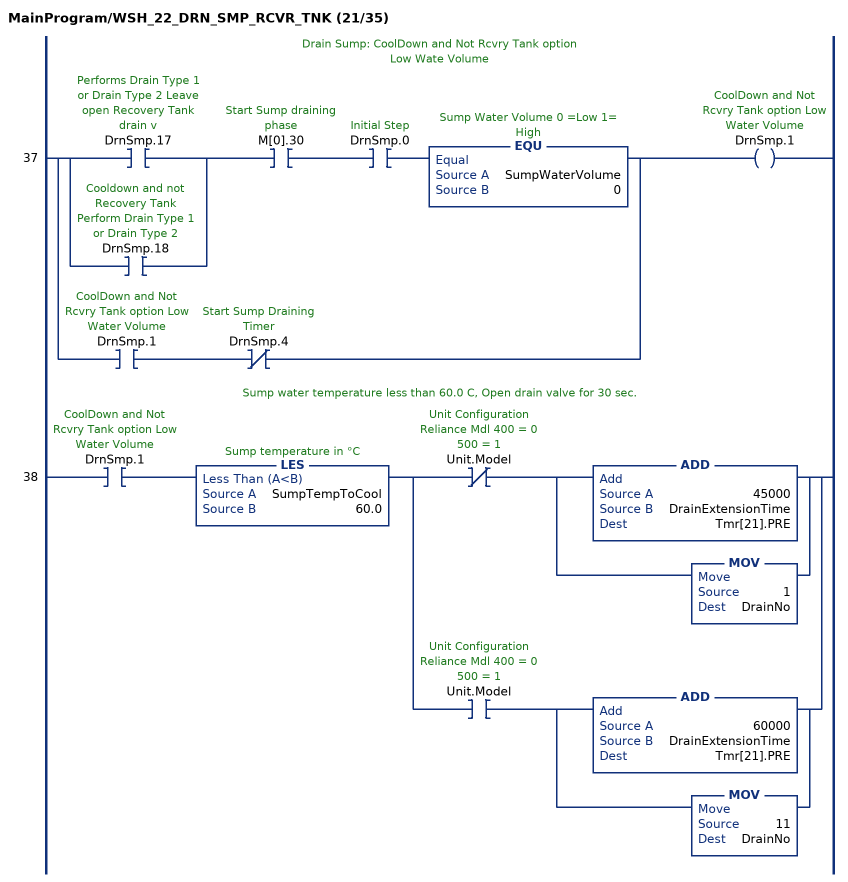
   // Drain Sump: CoolDown and Not Rcvry Tank option
   // Low Wate Volume
   37: [[XIC(DrnSmp.17) ,XIC(DrnSmp.18) ] XIC(M[0].30) XIC(DrnSmp.0) EQU(SumpWaterVolume,0) ,XIC(DrnSmp.1) XIO(DrnSmp.4) ]OTE(DrnSmp.1);
   // Sump water temperature less than 60.0 C, Open drain valve for 30 sec.
   38: XIC(DrnSmp.1)LES(SumpTempToCool,60.0)[XIO(Unit.Model) [ADD(45000,DrainExtensionTime,Tmr[21].PRE) ,MOV(1,DrainNo) ] ,XIC(Unit.Model) [ADD(60000,DrainExtensionTime,Tmr[21].PRE) ,MOV(11,DrainNo) ] ];
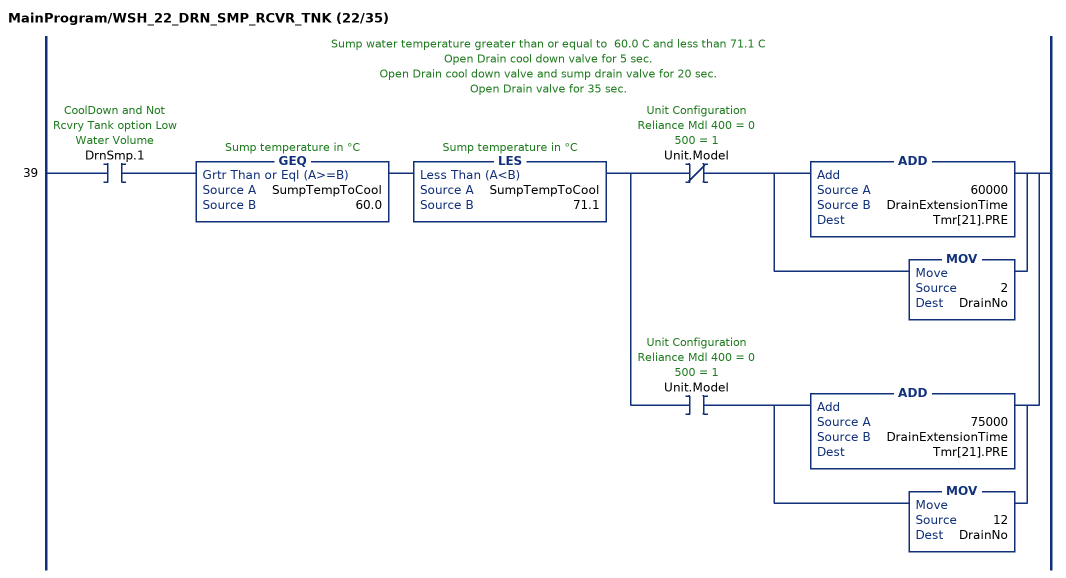
   // Sump water temperature greater than or equal to  60.0 C and less than 71.1 C
   // Open Drain cool down valve for 5 sec.
   // Open Drain cool down valve and sump drain valve for 20 sec.
   // Open Drain valve for 35 sec.
   39: XIC(DrnSmp.1)GEQ(SumpTempToCool,60.0)LES(SumpTempToCool,71.1)[XIO(Unit.Model) [ADD(60000,DrainExtensionTime,Tmr[21].PRE) ,MOV(2,DrainNo) ] ,XIC(Unit.Model) [ADD(75000,DrainExtensionTime,Tmr[21].PRE) ,MOV(12,DrainNo) ] ];
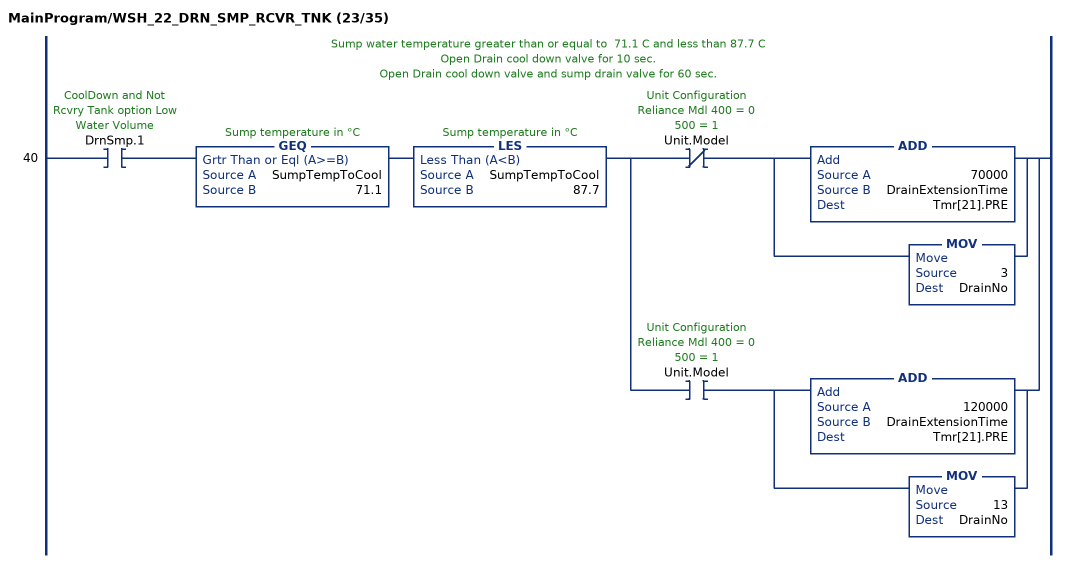
   // Sump water temperature greater than or equal to  71.1 C and less than 87.7 C
   // Open Drain cool down valve for 10 sec.
   // Open Drain cool down valve and sump drain valve for 60 sec.
   40: XIC(DrnSmp.1)GEQ(SumpTempToCool,71.1)LES(SumpTempToCool,87.7)[XIO(Unit.Model) [ADD(70000,DrainExtensionTime,Tmr[21].PRE) ,MOV(3,DrainNo) ] ,XIC(Unit.Model) [ADD(120000,DrainExtensionTime,Tmr[21].PRE) ,MOV(13,DrainNo) ] ];
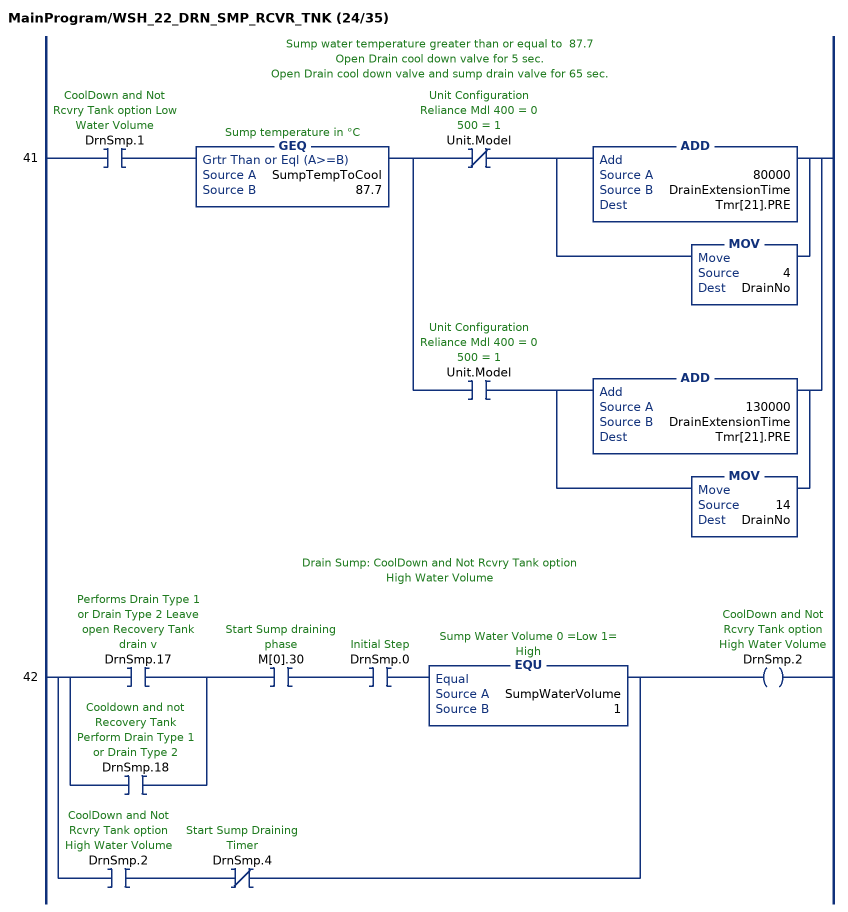
   // Sump water temperature greater than or equal to  87.7
   // Open Drain cool down valve for 5 sec.
   // Open Drain cool down valve and sump drain valve for 65 sec.
   41: XIC(DrnSmp.1)GEQ(SumpTempToCool,87.7)[XIO(Unit.Model) [ADD(80000,DrainExtensionTime,Tmr[21].PRE) ,MOV(4,DrainNo) ] ,XIC(Unit.Model) [ADD(130000,DrainExtensionTime,Tmr[21].PRE) ,MOV(14,DrainNo) ] ];
   // Drain Sump: CoolDown and Not Rcvry Tank option
   // High Water Volume
   42: [[XIC(DrnSmp.17) ,XIC(DrnSmp.18) ] XIC(M[0].30) XIC(DrnSmp.0) EQU(SumpWaterVolume,1) ,XIC(DrnSmp.2) XIO(DrnSmp.4) ]OTE(DrnSmp.2);
